// TIA Portal V20 export
// export: Created 2026-10-20T18:55:02.7661486Z, ExportSetting None, DisplayName Totally Integrated Automation Portal, DisplayVersion V20 Update 6, DisplayName TIA Portal Openness, DisplayVersion V20 Update 6, DisplayName TIA Portal Version Control Interface, DisplayVersion V20 Update 6, DisplayName SINAMICS Startdrive Advanced, DisplayVersion V20 SP1, DisplayName SINAMICS Startdrive G130, G150, S120, S150, SINAMICS MV, G220, S200, S210, DisplayVersion V20 SP1, DisplayName SINAMICS Startdrive G110M, G120, G120C, G120D, G120P, G115D, DisplayVersion V20 SP1, DisplayName STEP 7 Professional, DisplayVersion V20 Update 6, DisplayName STEP 7 Safety, DisplayVersion V20 Update 2, DisplayName WinCC Basic/Comfort/Advanced, DisplayVersion V20 Update 6, DisplayName WinCC Unified, DisplayVersion V20 Update 6
VAR_GLOBAL   // PLC tag table "IO_Turck_3"
   "Light_Front_1_1_Direction(3)" AT %QB837 : Byte;   // Last byte - 18
   "Light_Front_1_Animation(3)" AT %QB855 : Byte;   // Last byte
   "Light_Front_1_Pulse_Pattern(3)" AT %QB847 : Byte;   // Last byte - 8
   "Light_Rear_1_Color2(3)" AT %QB909 : Byte;   // Last byte - 10
   "Light_Front_1_Intensity2(3)" AT %QB843 : Byte;   // Last byte - 12
   "Light_Front_1_Bounce_Style(3)" AT %QB841 : Byte;   // Last byte - 14
   "Light_Rear_1_Color1(3)" AT %QB917 : Byte;   // Last byte - 2
   "Light_Front_1_Percent_Width1(3)" AT %QB839 : Byte;   // Last byte - 16
   "Light_Front_1_Intensity1(3)" AT %QB851 : Byte;   // Last byte - 4
   "Light_Rear_1_Intensity2(3)" AT %QB907 : Byte;   // Last byte - 12
   "Light_Rear_1_Pulse_Pattern(3)" AT %QB911 : Byte;   // Last byte - 8
   "Light_Rear_1_Animation(3)" AT %QB919 : Byte;   // Last byte
   "Light_Front_1_Speed(3)" AT %QB849 : Byte;   // Last byte - 6
   "Light_Rear_1_Direction(3)" AT %QB901 : Byte;   // Last byte - 18
   "Light_Rear_1_Percent_Width1(3)" AT %QB903 : Byte;   // Last byte - 16
   "Light_Rear_1_Intensity1(3)" AT %QB915 : Byte;   // Last byte - 4
   "Light_Rear_1_Bounce_Style(3)" AT %QB905 : Byte;   // Last byte - 14
   "Light_Rear_1_Speed(3)" AT %QB913 : Byte;   // Last byte - 6
   "Light_Front_1_Color1(3)" AT %QB853 : Byte;   // Last byte - 2
   "Light_Front_1_Color2(3)" AT %QB845 : Byte;   // Last byte - 10
END_VAR
